Fanuc KAREL source: KO00036.KL

PROGRAM KO00036
%NOLOCKGROUP
%ENVIRONMENT MIR
VAR
  P1: POSITION
  P2: POSITION
  F: BOOLEAN
  OUT: JOINTPOS
BEGIN
  F = TRUE
  OUT = MIRROR(P1, P2, F)
END KO00036
